Fanuc KAREL source: KT00886.KL

PROGRAM KT00886
%NOLOCKGROUP
VAR
  H1: ARRAY[2] OF SHORT
  H2: ARRAY[2] OF SHORT
  OUT: INTEGER
BEGIN
  H1[1] = 2
  H2[1] = 3
  H1[1] = 2
  H2[1] = 3
  OUT = ATAN2(H1[1], H1[1])
END KT00886
